RESOURCE RES0 : EMB_RES_ECO
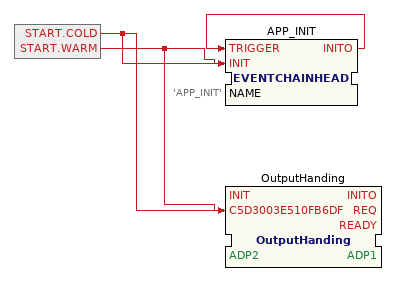
  FBS
    OutputHanding : OutputHanding;
    APP_INIT : EVENTCHAINHEAD(NAME := 'APP_INIT');
  END_FBS
  EVENT_CONNECTIONS
    APP_INIT.INITO TO APP_INIT.TRIGGER;
    START.COLD TO APP_INIT.INIT;
    START.WARM TO APP_INIT.INIT;
    START.COLD TO OutputHanding.C5D3003E510FB6DF;
    START.WARM TO OutputHanding.C5D3003E510FB6DF;
  END_CONNECTIONS
END_RESOURCE
